Staubli VAL3: logMoveMsgJ.pgx

program logMoveMsgJ(jointRx x_jPoint, tool x_tTool, mdesc x_mSpeed, num x_nMoveId, bool x_bExact)
  local string l_sCode
begin

  //
  if nRecIndex<200
    // j
    setMutex(bPushToStack)
    jPointRec[nRecIndex,1]=x_jPoint
    trToolRec[nRecIndex]=x_tTool.trsf
    mSpeedRec[nRecIndex]=x_mSpeed
    nMoveIdRec[nRecIndex]=x_nMoveId
    bExact[nRecIndex]=x_bExact
    nMoveTypeRec[nRecIndex]=2
    //logMsg("record moveJ."+toString("",nMoveIdRec[nRecIndex]))
    nRecIndex=nRecIndex+1
    bPushToStack=false
  else
    //popUpMsg("记录点数超过容量.")
  endIf

end
